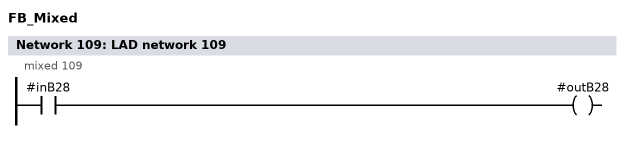
   RUNG wire#powerrail
      Contact( #inB28 )
      Coil( #outB28 )
   END_RUNG
   // the same network as SCL:
   #outB28 := #inB28;
END_REGION

REGION Network 110 (FBD): FBD network 110
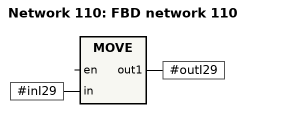
   #outI29 := #inI29;
END_REGION

REGION Network 111 (SCL): SCL network 111
   #tI10 := #inI30 + #cI20;
           IF #inB30 THEN
               #outR10 := #inR10 * 2.0;
           END_IF;
END_REGION

REGION Network 112: LAD network 112
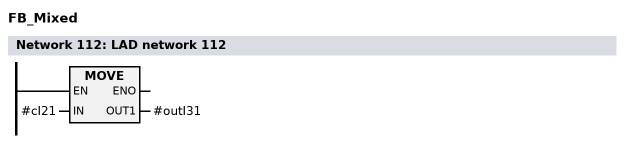
   RUNG wire#powerrail
      Move(in := #cI21, out1 => #outI31)
   END_RUNG
   // the same network as SCL:
   #outI31 := #cI21;
END_REGION

REGION Network 113 (FBD): FBD network 113
   // mixed 113
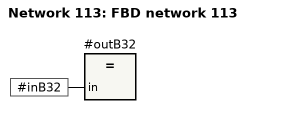
   #outB32 := #inB32;
END_REGION

REGION Network 114 (SCL): SCL network 114
   #tI13 := #inI33 + #cI23;
           IF #inB33 THEN
               #outR13 := #inR13 * 2.0;
           END_IF;
END_REGION

REGION Network 115: LAD network 115
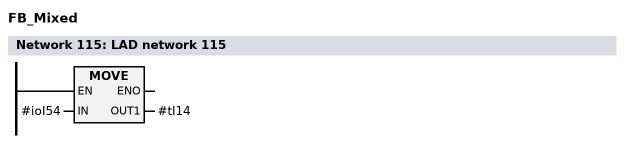
   RUNG wire#powerrail
      Move(in := #ioI54, out1 => #tI14)
   END_RUNG
   // the same network as SCL:
   #tI14 := #ioI54;
END_REGION

REGION Network 116 (FBD): FBD network 116
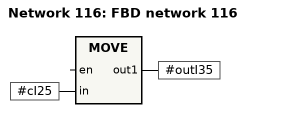
   #outI35 := #cI25;
END_REGION

REGION Network 117 (SCL): SCL network 117
   // mixed 117
   #tI16 := #inI36 + #cI26;
           IF #inB36 THEN
               #outR16 := #inR16 * 2.0;
           END_IF;
END_REGION

REGION Network 118: LAD network 118
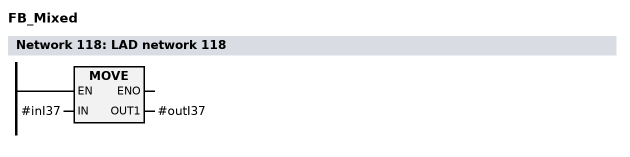
   RUNG wire#powerrail
      Move(in := #inI37, out1 => #outI37)
   END_RUNG
   // the same network as SCL:
   #outI37 := #inI37;
END_REGION

REGION Network 119 (FBD): FBD network 119
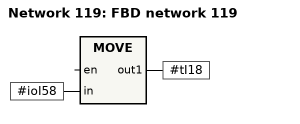
   #tI18 := #ioI58;
END_REGION

REGION Network 120 (SCL): SCL network 120
   #tI19 := #inI39 + #cI29;
           IF #inB39 THEN
               #outR19 := #inR19 * 2.0;
           END_IF;
END_REGION
END_FUNCTION_BLOCK

FUNCTION_BLOCK "FB_BigLad"   // FB14, LAD
{ S7_Optimized_Access := 'TRUE' }
VERSION : 0.1
   VAR_INPUT
      inB0 : Bool;   // input bit 0
      inB1 : Bool;
      inB2 : Bool;
      inB3 : Bool;
      inB4 : Bool;
      inB5 : Bool;
      inB6 : Bool;
      inB7 : Bool;
      inB8 : Bool;
      inB9 : Bool;
      inB10 : Bool;   // input bit 10
      inB11 : Bool;
      inB12 : Bool;
      inB13 : Bool;
      inB14 : Bool;
      inB15 : Bool;
      inB16 : Bool;
      inB17 : Bool;
      inB18 : Bool;
      inB19 : Bool;
      inB20 : Bool;   // input bit 20
      inB21 : Bool;
      inB22 : Bool;
      inB23 : Bool;
      inB24 : Bool;
      inB25 : Bool;
      inB26 : Bool;
      inB27 : Bool;
      inB28 : Bool;
      inB29 : Bool;
      inB30 : Bool;   // input bit 30
      inB31 : Bool;
      inB32 : Bool;
      inB33 : Bool;
      inB34 : Bool;
      inB35 : Bool;
      inB36 : Bool;
      inB37 : Bool;
      inB38 : Bool;
      inB39 : Bool;
      inI0 : Int;
      inI1 : Int;
      inI2 : Int;
      inI3 : Int;
      inI4 : Int;
      inI5 : Int;
      inI6 : Int;
      inI7 : Int;
      inI8 : Int;
      inI9 : Int;
      inI10 : Int;
      inI11 : Int;
      inI12 : Int;
      inI13 : Int;
      inI14 : Int;
      inI15 : Int;
      inI16 : Int;
      inI17 : Int;
      inI18 : Int;
      inI19 : Int;
      inI20 : Int;
      inI21 : Int;
      inI22 : Int;
      inI23 : Int;
      inI24 : Int;
      inI25 : Int;
      inI26 : Int;
      inI27 : Int;
      inI28 : Int;
      inI29 : Int;
      inI30 : Int;
      inI31 : Int;
      inI32 : Int;
      inI33 : Int;
      inI34 : Int;
      inI35 : Int;
      inI36 : Int;
      inI37 : Int;
      inI38 : Int;
      inI39 : Int;
      inR0 : Real;
      inR1 : Real;
      inR2 : Real;
      inR3 : Real;
      inR4 : Real;
      inR5 : Real;
      inR6 : Real;
      inR7 : Real;
      inR8 : Real;
      inR9 : Real;
      inR10 : Real;
      inR11 : Real;
      inR12 : Real;
      inR13 : Real;
      inR14 : Real;
      inR15 : Real;
      inR16 : Real;
      inR17 : Real;
      inR18 : Real;
      inR19 : Real;
      inD0 : DInt;
      inD1 : DInt;
      inD2 : DInt;
      inD3 : DInt;
      inD4 : DInt;
      inD5 : DInt;
      inD6 : DInt;
      inD7 : DInt;
      inD8 : DInt;
      inD9 : DInt;
      inD10 : DInt;
      inD11 : DInt;
      inD12 : DInt;
      inD13 : DInt;
      inD14 : DInt;
      inD15 : DInt;
      inD16 : DInt;
      inD17 : DInt;
      inD18 : DInt;
      inD19 : DInt;
      inArr : Array[0..99] of Int;   // input array
      inStr : String[40];
      inSt : Struct
         x : Int;
         y : Real;
         z : Bool;
      END_STRUCT;
   END_VAR
   VAR_OUTPUT
      outB0 : Bool;
      outB1 : Bool;
      outB2 : Bool;
      outB3 : Bool;
      outB4 : Bool;
      outB5 : Bool;
      outB6 : Bool;
      outB7 : Bool;
      outB8 : Bool;
      outB9 : Bool;
      outB10 : Bool;
      outB11 : Bool;
      outB12 : Bool;
      outB13 : Bool;
      outB14 : Bool;
      outB15 : Bool;
      outB16 : Bool;
      outB17 : Bool;
      outB18 : Bool;
      outB19 : Bool;
      outB20 : Bool;
      outB21 : Bool;
      outB22 : Bool;
      outB23 : Bool;
      outB24 : Bool;
      outB25 : Bool;
      outB26 : Bool;
      outB27 : Bool;
      outB28 : Bool;
      outB29 : Bool;
      outB30 : Bool;
      outB31 : Bool;
      outB32 : Bool;
      outB33 : Bool;
      outB34 : Bool;
      outB35 : Bool;
      outB36 : Bool;
      outB37 : Bool;
      outB38 : Bool;
      outB39 : Bool;
      outI0 : Int;   // output int 0
      outI1 : Int;
      outI2 : Int;
      outI3 : Int;
      outI4 : Int;
      outI5 : Int;
      outI6 : Int;
      outI7 : Int;
      outI8 : Int;
      outI9 : Int;
      outI10 : Int;   // output int 10
      outI11 : Int;
      outI12 : Int;
      outI13 : Int;
      outI14 : Int;
      outI15 : Int;
      outI16 : Int;
      outI17 : Int;
      outI18 : Int;
      outI19 : Int;
      outI20 : Int;   // output int 20
      outI21 : Int;
      outI22 : Int;
      outI23 : Int;
      outI24 : Int;
      outI25 : Int;
      outI26 : Int;
      outI27 : Int;
      outI28 : Int;
      outI29 : Int;
      outI30 : Int;   // output int 30
      outI31 : Int;
      outI32 : Int;
      outI33 : Int;
      outI34 : Int;
      outI35 : Int;
      outI36 : Int;
      outI37 : Int;
      outI38 : Int;
      outI39 : Int;
      outR0 : Real;
      outR1 : Real;
      outR2 : Real;
      outR3 : Real;
      outR4 : Real;
      outR5 : Real;
      outR6 : Real;
      outR7 : Real;
      outR8 : Real;
      outR9 : Real;
      outR10 : Real;
      outR11 : Real;
      outR12 : Real;
      outR13 : Real;
      outR14 : Real;
      outR15 : Real;
      outR16 : Real;
      outR17 : Real;
      outR18 : Real;
      outR19 : Real;
      outD0 : DInt;
      outD1 : DInt;
      outD2 : DInt;
      outD3 : DInt;
      outD4 : DInt;
      outD5 : DInt;
      outD6 : DInt;
      outD7 : DInt;
      outD8 : DInt;
      outD9 : DInt;
      outD10 : DInt;
      outD11 : DInt;
      outD12 : DInt;
      outD13 : DInt;
      outD14 : DInt;
      outD15 : DInt;
      outD16 : DInt;
      outD17 : DInt;
      outD18 : DInt;
      outD19 : DInt;
   END_VAR
   VAR_IN_OUT
      ioI0 : Int;
      ioI1 : Int;
      ioI2 : Int;
      ioI3 : Int;
      ioI4 : Int;
      ioI5 : Int;
      ioI6 : Int;
      ioI7 : Int;
      ioI8 : Int;
      ioI9 : Int;
      ioI10 : Int;
      ioI11 : Int;
      ioI12 : Int;
      ioI13 : Int;
      ioI14 : Int;
      ioI15 : Int;
      ioI16 : Int;
      ioI17 : Int;
      ioI18 : Int;
      ioI19 : Int;
      ioI20 : Int;
      ioI21 : Int;
      ioI22 : Int;
      ioI23 : Int;
      ioI24 : Int;
      ioI25 : Int;
      ioI26 : Int;
      ioI27 : Int;
      ioI28 : Int;
      ioI29 : Int;
      ioI30 : Int;
      ioI31 : Int;
      ioI32 : Int;
      ioI33 : Int;
      ioI34 : Int;
      ioI35 : Int;
      ioI36 : Int;
      ioI37 : Int;
      ioI38 : Int;
      ioI39 : Int;
      ioI40 : Int;
      ioI41 : Int;
      ioI42 : Int;
      ioI43 : Int;
      ioI44 : Int;
      ioI45 : Int;
      ioI46 : Int;
      ioI47 : Int;
      ioI48 : Int;
      ioI49 : Int;
      ioI50 : Int;
      ioI51 : Int;
      ioI52 : Int;
      ioI53 : Int;
      ioI54 : Int;
      ioI55 : Int;
      ioI56 : Int;
      ioI57 : Int;
      ioI58 : Int;
      ioI59 : Int;
   END_VAR
   VAR
      stI0 : Int := 0;   // static 0
      stI1 : Int;
      stI2 : Int;
      stI3 : Int;
      stI4 : Int;
      stI5 : Int;
      stI6 : Int;
      stI7 : Int := 7;
      stI8 : Int;
      stI9 : Int;
      stI10 : Int;
      stI11 : Int;
      stI12 : Int;
      stI13 : Int;
      stI14 : Int := 14;
      stI15 : Int;
      stI16 : Int;
      stI17 : Int;
      stI18 : Int;
      stI19 : Int;
      stI20 : Int;
      stI21 : Int := 21;
      stI22 : Int;
      stI23 : Int;
      stI24 : Int;
      stI25 : Int;   // static 25
      stI26 : Int;
      stI27 : Int;
      stI28 : Int := 28;
      stI29 : Int;
      stI30 : Int;
      stI31 : Int;
      stI32 : Int;
      stI33 : Int;
      stI34 : Int;
      stI35 : Int := 35;
      stI36 : Int;
      stI37 : Int;
      stI38 : Int;
      stI39 : Int;
      stI40 : Int;
      stI41 : Int;
      stI42 : Int := 42;
      stI43 : Int;
      stI44 : Int;
      stI45 : Int;
      stI46 : Int;
      stI47 : Int;
      stI48 : Int;
      stI49 : Int := 49;
      stI50 : Int;   // static 50
      stI51 : Int;
      stI52 : Int;
      stI53 : Int;
      stI54 : Int;
      stI55 : Int;
      stI56 : Int := 56;
      stI57 : Int;
      stI58 : Int;
      stI59 : Int;
      stI60 : Int;
      stI61 : Int;
      stI62 : Int;
      stI63 : Int := 63;
      stI64 : Int;
      stI65 : Int;
      stI66 : Int;
      stI67 : Int;
      stI68 : Int;
      stI69 : Int;
      stI70 : Int := 70;
      stI71 : Int;
      stI72 : Int;
      stI73 : Int;
      stI74 : Int;
      stI75 : Int;   // static 75
      stI76 : Int;
      stI77 : Int := 77;
      stI78 : Int;
      stI79 : Int;
      stI80 : Int;
      stI81 : Int;
      stI82 : Int;
      stI83 : Int;
      stI84 : Int := 84;
      stI85 : Int;
      stI86 : Int;
      stI87 : Int;
      stI88 : Int;
      stI89 : Int;
      stI90 : Int;
      stI91 : Int := 91;
      stI92 : Int;
      stI93 : Int;
      stI94 : Int;
      stI95 : Int;
      stI96 : Int;
      stI97 : Int;
      stI98 : Int := 98;
      stI99 : Int;
      stI100 : Int;   // static 100
      stI101 : Int;
      stI102 : Int;
      stI103 : Int;
      stI104 : Int;
      stI105 : Int := 105;
      stI106 : Int;
      stI107 : Int;
      stI108 : Int;
      stI109 : Int;
      stI110 : Int;
      stI111 : Int;
      stI112 : Int := 112;
      stI113 : Int;
      stI114 : Int;
      stI115 : Int;
      stI116 : Int;
      stI117 : Int;
      stI118 : Int;
      stI119 : Int := 119;
      stI120 : Int;
      stI121 : Int;
      stI122 : Int;
      stI123 : Int;
      stI124 : Int;
      stI125 : Int;   // static 125
      stI126 : Int := 126;
      stI127 : Int;
      stI128 : Int;
      stI129 : Int;
      stI130 : Int;
      stI131 : Int;
      stI132 : Int;
      stI133 : Int := 133;
      stI134 : Int;
      stI135 : Int;
      stI136 : Int;
      stI137 : Int;
      stI138 : Int;
      stI139 : Int;
      stI140 : Int := 140;
      stI141 : Int;
      stI142 : Int;
      stI143 : Int;
      stI144 : Int;
      stI145 : Int;
      stI146 : Int;
      stI147 : Int := 147;
      stI148 : Int;
      stI149 : Int;
      stI150 : Int;   // static 150
      stI151 : Int;
      stI152 : Int;
      stI153 : Int;
      stI154 : Int := 154;
      stI155 : Int;
      stI156 : Int;
      stI157 : Int;
      stI158 : Int;
      stI159 : Int;
      stI160 : Int;
      stI161 : Int := 161;
      stI162 : Int;
      stI163 : Int;
      stI164 : Int;
      stI165 : Int;
      stI166 : Int;
      stI167 : Int;
      stI168 : Int := 168;
      stI169 : Int;
      stI170 : Int;
      stI171 : Int;
      stI172 : Int;
      stI173 : Int;
      stI174 : Int;
      stI175 : Int := 175;   // static 175
      stI176 : Int;
      stI177 : Int;
      stI178 : Int;
      stI179 : Int;
      stI180 : Int;
      stI181 : Int;
      stI182 : Int := 182;
      stI183 : Int;
      stI184 : Int;
      stI185 : Int;
      stI186 : Int;
      stI187 : Int;
      stI188 : Int;
      stI189 : Int := 189;
      stI190 : Int;
      stI191 : Int;
      stI192 : Int;
      stI193 : Int;
      stI194 : Int;
      stI195 : Int;
      stI196 : Int := 196;
      stI197 : Int;
      stI198 : Int;
      stI199 : Int;
      stB0 : Bool := TRUE;
      stB1 : Bool;
      stB2 : Bool;
      stB3 : Bool := TRUE;
      stB4 : Bool;
      stB5 : Bool;
      stB6 : Bool := TRUE;
      stB7 : Bool;
      stB8 : Bool;
      stB9 : Bool := TRUE;
      stB10 : Bool;
      stB11 : Bool;
      stB12 : Bool := TRUE;
      stB13 : Bool;
      stB14 : Bool;
      stB15 : Bool := TRUE;
      stB16 : Bool;
      stB17 : Bool;
      stB18 : Bool := TRUE;
      stB19 : Bool;
      stB20 : Bool;
      stB21 : Bool := TRUE;
      stB22 : Bool;
      stB23 : Bool;
      stB24 : Bool := TRUE;
      stB25 : Bool;
      stB26 : Bool;
      stB27 : Bool := TRUE;
      stB28 : Bool;
      stB29 : Bool;
      stB30 : Bool := TRUE;
      stB31 : Bool;
      stB32 : Bool;
      stB33 : Bool := TRUE;
      stB34 : Bool;
      stB35 : Bool;
      stB36 : Bool := TRUE;
      stB37 : Bool;
      stB38 : Bool;
      stB39 : Bool := TRUE;
      stB40 : Bool;
      stB41 : Bool;
      stB42 : Bool := TRUE;
      stB43 : Bool;
      stB44 : Bool;
      stB45 : Bool := TRUE;
      stB46 : Bool;
      stB47 : Bool;
      stB48 : Bool := TRUE;
      stB49 : Bool;
      stB50 : Bool;
      stB51 : Bool := TRUE;
      stB52 : Bool;
      stB53 : Bool;
      stB54 : Bool := TRUE;
      stB55 : Bool;
      stB56 : Bool;
      stB57 : Bool := TRUE;
      stB58 : Bool;
      stB59 : Bool;
      stB60 : Bool := TRUE;
      stB61 : Bool;
      stB62 : Bool;
      stB63 : Bool := TRUE;
      stB64 : Bool;
      stB65 : Bool;
      stB66 : Bool := TRUE;
      stB67 : Bool;
      stB68 : Bool;
      stB69 : Bool := TRUE;
      stB70 : Bool;
      stB71 : Bool;
      stB72 : Bool := TRUE;
      stB73 : Bool;
      stB74 : Bool;
      stB75 : Bool := TRUE;
      stB76 : Bool;
      stB77 : Bool;
      stB78 : Bool := TRUE;
      stB79 : Bool;
      stB80 : Bool;
      stB81 : Bool := TRUE;
      stB82 : Bool;
      stB83 : Bool;
      stB84 : Bool := TRUE;
      stB85 : Bool;
      stB86 : Bool;
      stB87 : Bool := TRUE;
      stB88 : Bool;
      stB89 : Bool;
      stB90 : Bool := TRUE;
      stB91 : Bool;
      stB92 : Bool;
      stB93 : Bool := TRUE;
      stB94 : Bool;
      stB95 : Bool;
      stB96 : Bool := TRUE;
      stB97 : Bool;
      stB98 : Bool;
      stB99 : Bool := TRUE;
      stArr : Array[1..10, 0..4] of Real;
      stSt : Struct
         "a" : Int;
         "b" : Array[0..3] of Bool;
         c : Time;
      END_STRUCT;
   END_VAR
   VAR_TEMP
      tI0 : Int;
      tI1 : Int;
      tI2 : Int;
      tI3 : Int;
      tI4 : Int;
      tI5 : Int;
      tI6 : Int;
      tI7 : Int;
      tI8 : Int;
      tI9 : Int;
      tI10 : Int;
      tI11 : Int;
      tI12 : Int;
      tI13 : Int;
      tI14 : Int;
      tI15 : Int;
      tI16 : Int;
      tI17 : Int;
      tI18 : Int;
      tI19 : Int;
      tI20 : Int;
      tI21 : Int;
      tI22 : Int;
      tI23 : Int;
      tI24 : Int;
      tI25 : Int;
      tI26 : Int;
      tI27 : Int;
      tI28 : Int;
      tI29 : Int;
      tI30 : Int;
      tI31 : Int;
      tI32 : Int;
      tI33 : Int;
      tI34 : Int;
      tI35 : Int;
      tI36 : Int;
      tI37 : Int;
      tI38 : Int;
      tI39 : Int;
      tI40 : Int;
      tI41 : Int;
      tI42 : Int;
      tI43 : Int;
      tI44 : Int;
      tI45 : Int;
      tI46 : Int;
      tI47 : Int;
      tI48 : Int;
      tI49 : Int;
      tI50 : Int;
      tI51 : Int;
      tI52 : Int;
      tI53 : Int;
      tI54 : Int;
      tI55 : Int;
      tI56 : Int;
      tI57 : Int;
      tI58 : Int;
      tI59 : Int;
      tI60 : Int;
      tI61 : Int;
      tI62 : Int;
      tI63 : Int;
      tI64 : Int;
      tI65 : Int;
      tI66 : Int;
      tI67 : Int;
      tI68 : Int;
      tI69 : Int;
      tI70 : Int;
      tI71 : Int;
      tI72 : Int;
      tI73 : Int;
      tI74 : Int;
      tI75 : Int;
      tI76 : Int;
      tI77 : Int;
      tI78 : Int;
      tI79 : Int;
      tI80 : Int;
      tI81 : Int;
      tI82 : Int;
      tI83 : Int;
      tI84 : Int;
      tI85 : Int;
      tI86 : Int;
      tI87 : Int;
      tI88 : Int;
      tI89 : Int;
      tI90 : Int;
      tI91 : Int;
      tI92 : Int;
      tI93 : Int;
      tI94 : Int;
      tI95 : Int;
      tI96 : Int;
      tI97 : Int;
      tI98 : Int;
      tI99 : Int;
      tR0 : Real;
      tR1 : Real;
      tR2 : Real;
      tR3 : Real;
      tR4 : Real;
      tR5 : Real;
      tR6 : Real;
      tR7 : Real;
      tR8 : Real;
      tR9 : Real;
      tR10 : Real;
      tR11 : Real;
      tR12 : Real;
      tR13 : Real;
      tR14 : Real;
      tR15 : Real;
      tR16 : Real;
      tR17 : Real;
      tR18 : Real;
      tR19 : Real;
      tR20 : Real;
      tR21 : Real;
      tR22 : Real;
      tR23 : Real;
      tR24 : Real;
      tR25 : Real;
      tR26 : Real;
      tR27 : Real;
      tR28 : Real;
      tR29 : Real;
      tR30 : Real;
      tR31 : Real;
      tR32 : Real;
      tR33 : Real;
      tR34 : Real;
      tR35 : Real;
      tR36 : Real;
      tR37 : Real;
      tR38 : Real;
      tR39 : Real;
      tR40 : Real;
      tR41 : Real;
      tR42 : Real;
      tR43 : Real;
      tR44 : Real;
      tR45 : Real;
      tR46 : Real;
      tR47 : Real;
      tR48 : Real;
      tR49 : Real;
   END_VAR
   VAR CONSTANT
      cI0 : Int := 0;
      cI1 : Int := 3;
      cI2 : Int := 6;
      cI3 : Int := 9;
      cI4 : Int := 12;
      cI5 : Int := 15;
      cI6 : Int := 18;
      cI7 : Int := 21;
      cI8 : Int := 24;
      cI9 : Int := 27;
      cI10 : Int := 30;
      cI11 : Int := 33;
      cI12 : Int := 36;
      cI13 : Int := 39;
      cI14 : Int := 42;
      cI15 : Int := 45;
      cI16 : Int := 48;
      cI17 : Int := 51;
      cI18 : Int := 54;
      cI19 : Int := 57;
      cI20 : Int := 60;
      cI21 : Int := 63;
      cI22 : Int := 66;
      cI23 : Int := 69;
      cI24 : Int := 72;
      cI25 : Int := 75;
      cI26 : Int := 78;
      cI27 : Int := 81;
      cI28 : Int := 84;
      cI29 : Int := 87;
   END_VAR
BEGIN

REGION Network 1: LAD network 1
   // comment of network 1
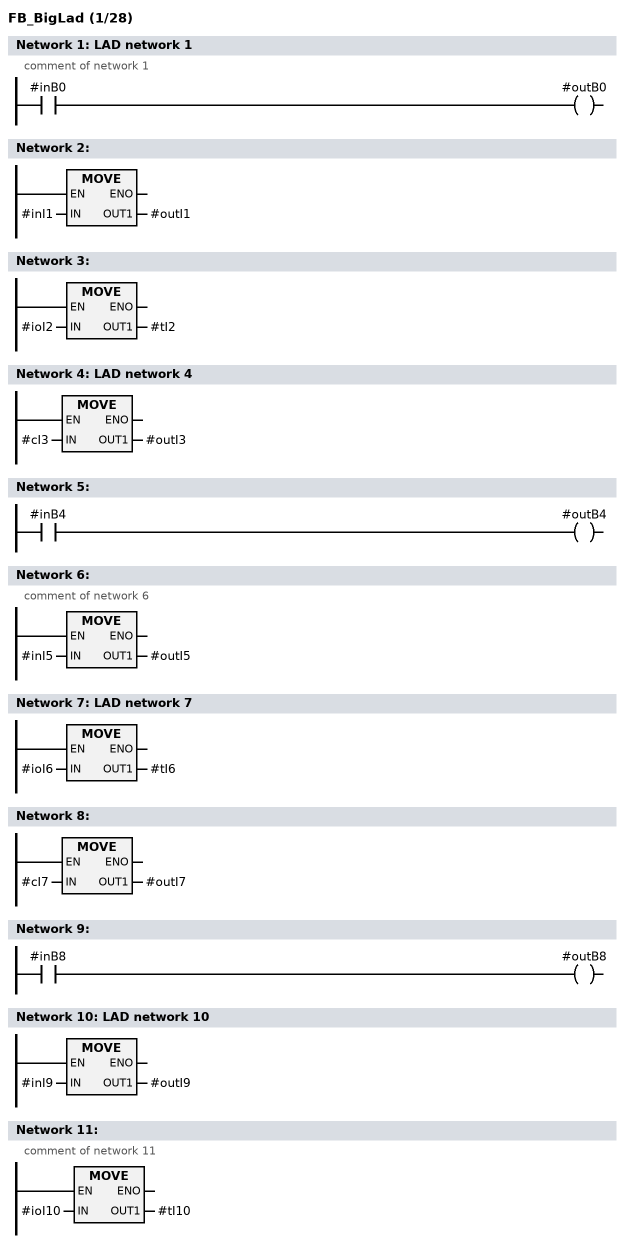
   RUNG wire#powerrail
      Contact( #inB0 )
      Coil( #outB0 )
   END_RUNG
   // the same network as SCL:
   #outB0 := #inB0;
END_REGION

REGION Network 2
   RUNG wire#powerrail
      Move(in := #inI1, out1 => #outI1)
   END_RUNG
   // the same network as SCL:
   #outI1 := #inI1;
END_REGION

REGION Network 3
   RUNG wire#powerrail
      Move(in := #ioI2, out1 => #tI2)
   END_RUNG
   // the same network as SCL:
   #tI2 := #ioI2;
END_REGION

REGION Network 4: LAD network 4
   RUNG wire#powerrail
      Move(in := #cI3, out1 => #outI3)
   END_RUNG
   // the same network as SCL:
   #outI3 := #cI3;
END_REGION

REGION Network 5
   RUNG wire#powerrail
      Contact( #inB4 )
      Coil( #outB4 )
   END_RUNG
   // the same network as SCL:
   #outB4 := #inB4;
END_REGION

REGION Network 6
   // comment of network 6
   RUNG wire#powerrail
      Move(in := #inI5, out1 => #outI5)
   END_RUNG
   // the same network as SCL:
   #outI5 := #inI5;
END_REGION

REGION Network 7: LAD network 7
   RUNG wire#powerrail
      Move(in := #ioI6, out1 => #tI6)
   END_RUNG
   // the same network as SCL:
   #tI6 := #ioI6;
END_REGION

REGION Network 8
   RUNG wire#powerrail
      Move(in := #cI7, out1 => #outI7)
   END_RUNG
   // the same network as SCL:
   #outI7 := #cI7;
END_REGION

REGION Network 9
   RUNG wire#powerrail
      Contact( #inB8 )
      Coil( #outB8 )
   END_RUNG
   // the same network as SCL:
   #outB8 := #inB8;
END_REGION

REGION Network 10: LAD network 10
   RUNG wire#powerrail
      Move(in := #inI9, out1 => #outI9)
   END_RUNG
   // the same network as SCL:
   #outI9 := #inI9;
END_REGION

REGION Network 11
   // comment of network 11
   RUNG wire#powerrail
      Move(in := #ioI10, out1 => #tI10)
   END_RUNG
   // the same network as SCL:
   #tI10 := #ioI10;
END_REGION

REGION Network 12
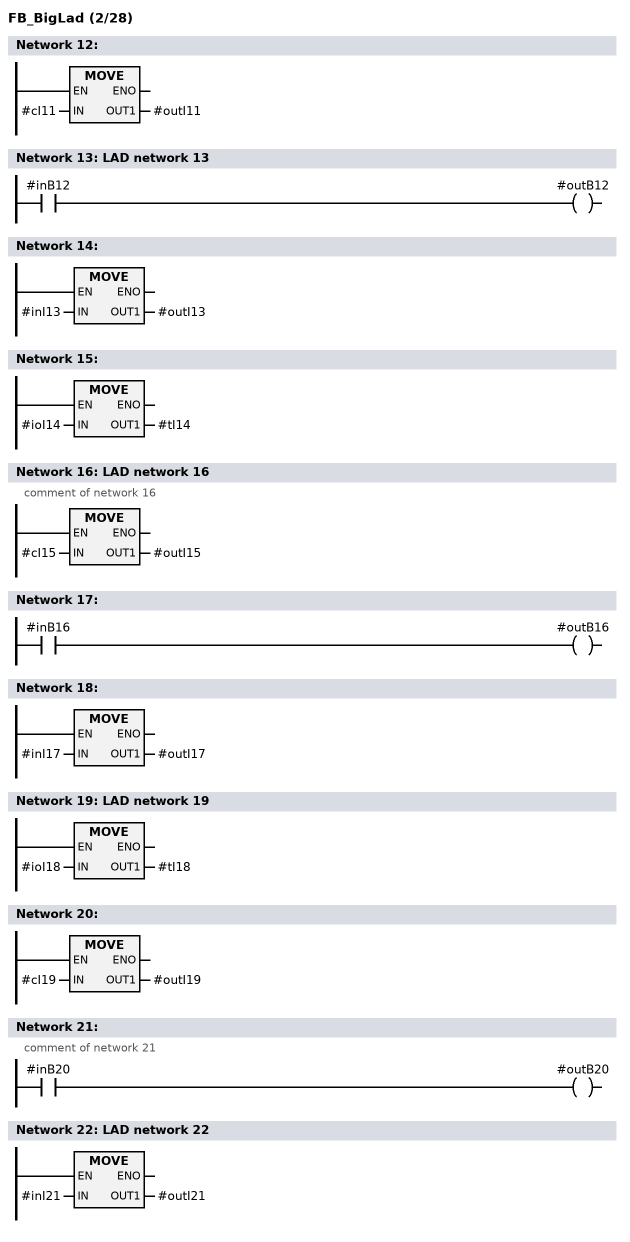
   RUNG wire#powerrail
      Move(in := #cI11, out1 => #outI11)
   END_RUNG
   // the same network as SCL:
   #outI11 := #cI11;
END_REGION

REGION Network 13: LAD network 13
   RUNG wire#powerrail
      Contact( #inB12 )
      Coil( #outB12 )
   END_RUNG
   // the same network as SCL:
   #outB12 := #inB12;
END_REGION

REGION Network 14
   RUNG wire#powerrail
      Move(in := #inI13, out1 => #outI13)
   END_RUNG
   // the same network as SCL:
   #outI13 := #inI13;
END_REGION

REGION Network 15
   RUNG wire#powerrail
      Move(in := #ioI14, out1 => #tI14)
   END_RUNG
   // the same network as SCL:
   #tI14 := #ioI14;
END_REGION

REGION Network 16: LAD network 16
   // comment of network 16
   RUNG wire#powerrail
      Move(in := #cI15, out1 => #outI15)
   END_RUNG
   // the same network as SCL:
   #outI15 := #cI15;
END_REGION

REGION Network 17
   RUNG wire#powerrail
      Contact( #inB16 )
      Coil( #outB16 )
   END_RUNG
   // the same network as SCL:
   #outB16 := #inB16;
END_REGION

REGION Network 18
   RUNG wire#powerrail
      Move(in := #inI17, out1 => #outI17)
   END_RUNG
   // the same network as SCL:
   #outI17 := #inI17;
END_REGION

REGION Network 19: LAD network 19
   RUNG wire#powerrail
      Move(in := #ioI18, out1 => #tI18)
   END_RUNG
   // the same network as SCL:
   #tI18 := #ioI18;
END_REGION

REGION Network 20
   RUNG wire#powerrail
      Move(in := #cI19, out1 => #outI19)
   END_RUNG
   // the same network as SCL:
   #outI19 := #cI19;
END_REGION

REGION Network 21
   // comment of network 21
   RUNG wire#powerrail
      Contact( #inB20 )
      Coil( #outB20 )
   END_RUNG
   // the same network as SCL:
   #outB20 := #inB20;
END_REGION

REGION Network 22: LAD network 22
   RUNG wire#powerrail
      Move(in := #inI21, out1 => #outI21)
   END_RUNG
   // the same network as SCL:
   #outI21 := #inI21;
END_REGION

REGION Network 23
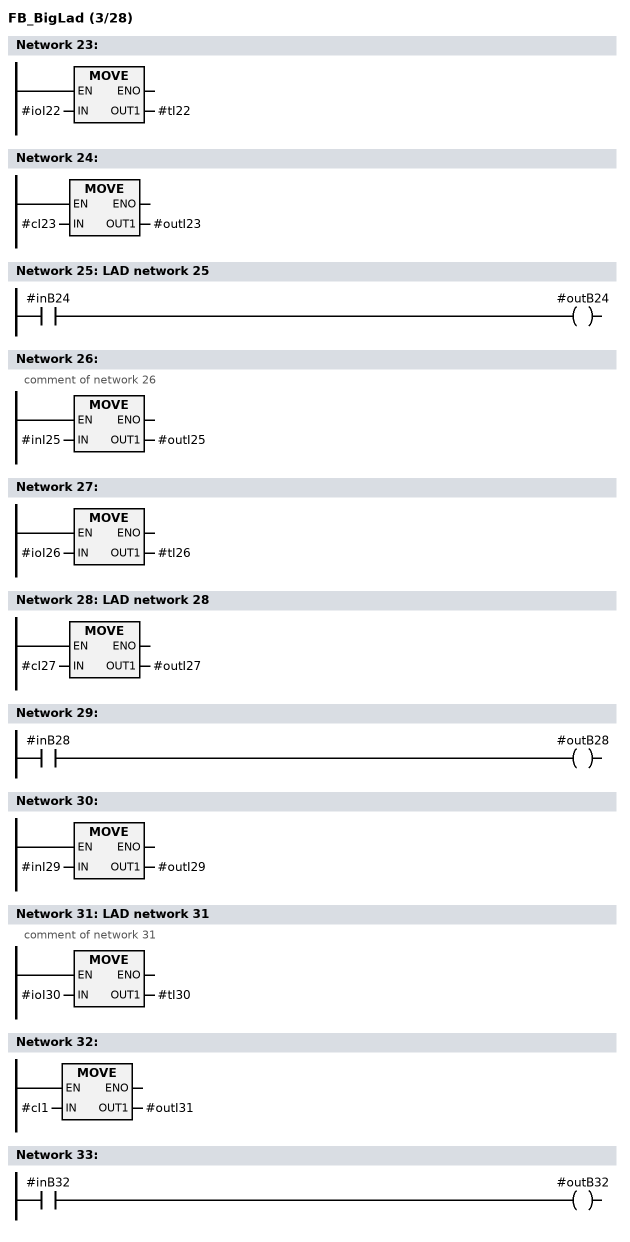
   RUNG wire#powerrail
      Move(in := #ioI22, out1 => #tI22)
   END_RUNG
   // the same network as SCL:
   #tI22 := #ioI22;
END_REGION

REGION Network 24
   RUNG wire#powerrail
      Move(in := #cI23, out1 => #outI23)
   END_RUNG
   // the same network as SCL:
   #outI23 := #cI23;
END_REGION

REGION Network 25: LAD network 25
   RUNG wire#powerrail
      Contact( #inB24 )
      Coil( #outB24 )
   END_RUNG
   // the same network as SCL:
   #outB24 := #inB24;
END_REGION

REGION Network 26
   // comment of network 26
   RUNG wire#powerrail
      Move(in := #inI25, out1 => #outI25)
   END_RUNG
   // the same network as SCL:
   #outI25 := #inI25;
END_REGION

REGION Network 27
   RUNG wire#powerrail
      Move(in := #ioI26, out1 => #tI26)
   END_RUNG
   // the same network as SCL:
   #tI26 := #ioI26;
END_REGION

REGION Network 28: LAD network 28
   RUNG wire#powerrail
      Move(in := #cI27, out1 => #outI27)
   END_RUNG
   // the same network as SCL:
   #outI27 := #cI27;
END_REGION

REGION Network 29
   RUNG wire#powerrail
      Contact( #inB28 )
      Coil( #outB28 )
   END_RUNG
   // the same network as SCL:
   #outB28 := #inB28;
END_REGION

REGION Network 30
   RUNG wire#powerrail
      Move(in := #inI29, out1 => #outI29)
   END_RUNG
   // the same network as SCL:
   #outI29 := #inI29;
END_REGION

REGION Network 31: LAD network 31
   // comment of network 31
   RUNG wire#powerrail
      Move(in := #ioI30, out1 => #tI30)
   END_RUNG
   // the same network as SCL:
   #tI30 := #ioI30;
END_REGION

REGION Network 32
   RUNG wire#powerrail
      Move(in := #cI1, out1 => #outI31)
   END_RUNG
   // the same network as SCL:
   #outI31 := #cI1;
END_REGION

REGION Network 33
   RUNG wire#powerrail
      Contact( #inB32 )
      Coil( #outB32 )
   END_RUNG
   // the same network as SCL:
   #outB32 := #inB32;
END_REGION

REGION Network 34: LAD network 34
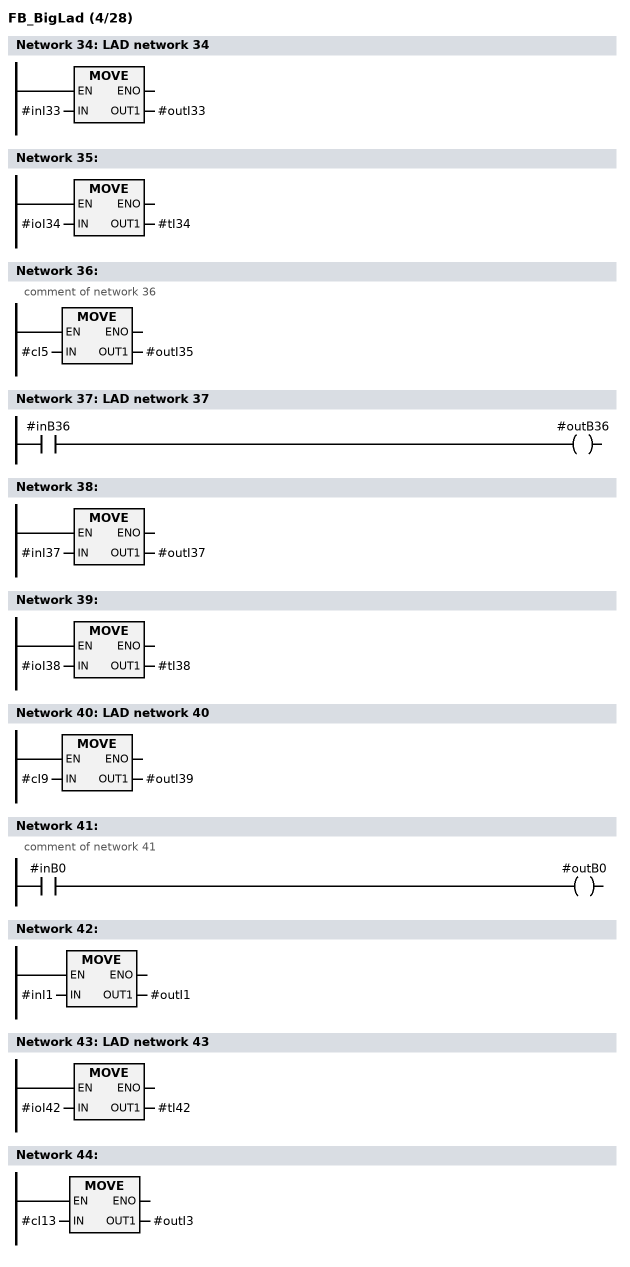
   RUNG wire#powerrail
      Move(in := #inI33, out1 => #outI33)
   END_RUNG
   // the same network as SCL:
   #outI33 := #inI33;
END_REGION

REGION Network 35
   RUNG wire#powerrail
      Move(in := #ioI34, out1 => #tI34)
   END_RUNG
   // the same network as SCL:
   #tI34 := #ioI34;
END_REGION

REGION Network 36
   // comment of network 36
   RUNG wire#powerrail
      Move(in := #cI5, out1 => #outI35)
   END_RUNG
   // the same network as SCL:
   #outI35 := #cI5;
END_REGION

REGION Network 37: LAD network 37
   RUNG wire#powerrail
      Contact( #inB36 )
      Coil( #outB36 )
   END_RUNG
   // the same network as SCL:
   #outB36 := #inB36;
END_REGION

REGION Network 38
   RUNG wire#powerrail
      Move(in := #inI37, out1 => #outI37)
   END_RUNG
   // the same network as SCL:
   #outI37 := #inI37;
END_REGION

REGION Network 39
   RUNG wire#powerrail
      Move(in := #ioI38, out1 => #tI38)
   END_RUNG
   // the same network as SCL:
   #tI38 := #ioI38;
END_REGION

REGION Network 40: LAD network 40
   RUNG wire#powerrail
      Move(in := #cI9, out1 => #outI39)
   END_RUNG
   // the same network as SCL:
   #outI39 := #cI9;
END_REGION

REGION Network 41
   // comment of network 41
   RUNG wire#powerrail
      Contact( #inB0 )
      Coil( #outB0 )
   END_RUNG
   // the same network as SCL:
   #outB0 := #inB0;
END_REGION

REGION Network 42
   RUNG wire#powerrail
      Move(in := #inI1, out1 => #outI1)
   END_RUNG
   // the same network as SCL:
   #outI1 := #inI1;
END_REGION

REGION Network 43: LAD network 43
   RUNG wire#powerrail
      Move(in := #ioI42, out1 => #tI42)
   END_RUNG
   // the same network as SCL:
   #tI42 := #ioI42;
END_REGION

REGION Network 44
   RUNG wire#powerrail
      Move(in := #cI13, out1 => #outI3)
   END_RUNG
   // the same network as SCL:
   #outI3 := #cI13;
END_REGION

REGION Network 45
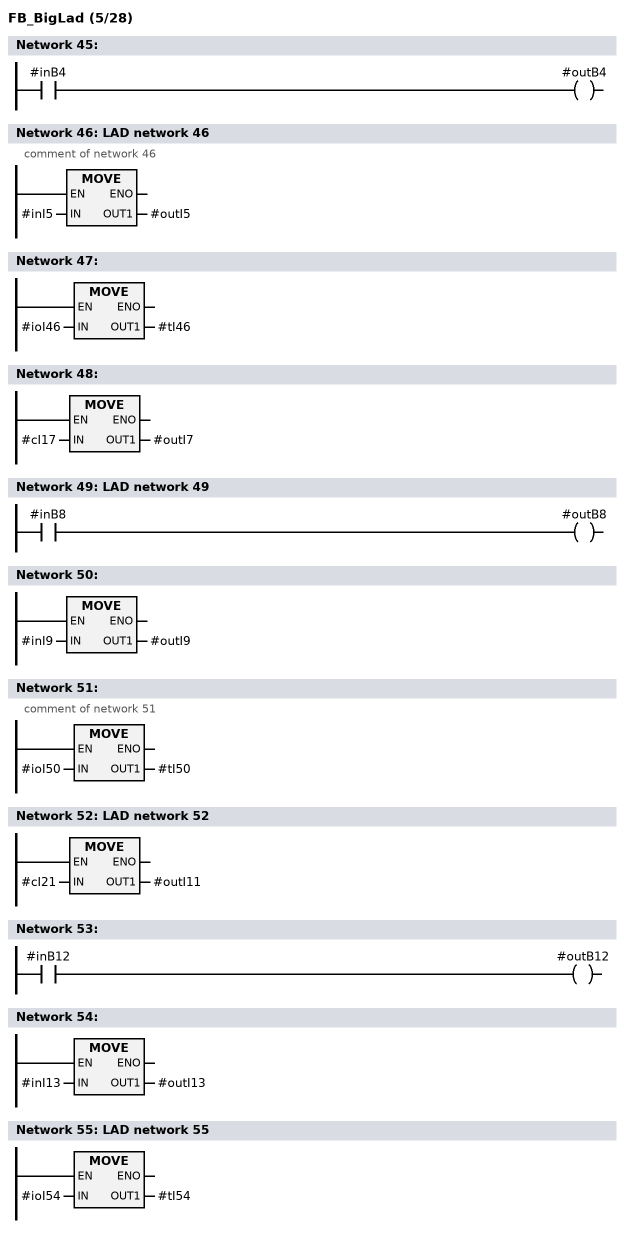
   RUNG wire#powerrail
      Contact( #inB4 )
      Coil( #outB4 )
   END_RUNG
   // the same network as SCL:
   #outB4 := #inB4;
END_REGION

REGION Network 46: LAD network 46
   // comment of network 46
   RUNG wire#powerrail
      Move(in := #inI5, out1 => #outI5)
   END_RUNG
   // the same network as SCL:
   #outI5 := #inI5;
END_REGION

REGION Network 47
   RUNG wire#powerrail
      Move(in := #ioI46, out1 => #tI46)
   END_RUNG
   // the same network as SCL:
   #tI46 := #ioI46;
END_REGION

REGION Network 48
   RUNG wire#powerrail
      Move(in := #cI17, out1 => #outI7)
   END_RUNG
   // the same network as SCL:
   #outI7 := #cI17;
END_REGION

REGION Network 49: LAD network 49
   RUNG wire#powerrail
      Contact( #inB8 )
      Coil( #outB8 )
   END_RUNG
   // the same network as SCL:
   #outB8 := #inB8;
END_REGION

REGION Network 50
   RUNG wire#powerrail
      Move(in := #inI9, out1 => #outI9)
   END_RUNG
   // the same network as SCL:
   #outI9 := #inI9;
END_REGION

REGION Network 51
   // comment of network 51
   RUNG wire#powerrail
      Move(in := #ioI50, out1 => #tI50)
   END_RUNG
   // the same network as SCL:
   #tI50 := #ioI50;
END_REGION

REGION Network 52: LAD network 52
   RUNG wire#powerrail
      Move(in := #cI21, out1 => #outI11)
   END_RUNG
   // the same network as SCL:
   #outI11 := #cI21;
END_REGION

REGION Network 53
   RUNG wire#powerrail
      Contact( #inB12 )
      Coil( #outB12 )
   END_RUNG
   // the same network as SCL:
   #outB12 := #inB12;
END_REGION

REGION Network 54
   RUNG wire#powerrail
      Move(in := #inI13, out1 => #outI13)
   END_RUNG
   // the same network as SCL:
   #outI13 := #inI13;
END_REGION

REGION Network 55: LAD network 55
   RUNG wire#powerrail
      Move(in := #ioI54, out1 => #tI54)
   END_RUNG
   // the same network as SCL:
   #tI54 := #ioI54;
END_REGION

REGION Network 56
   // comment of network 56
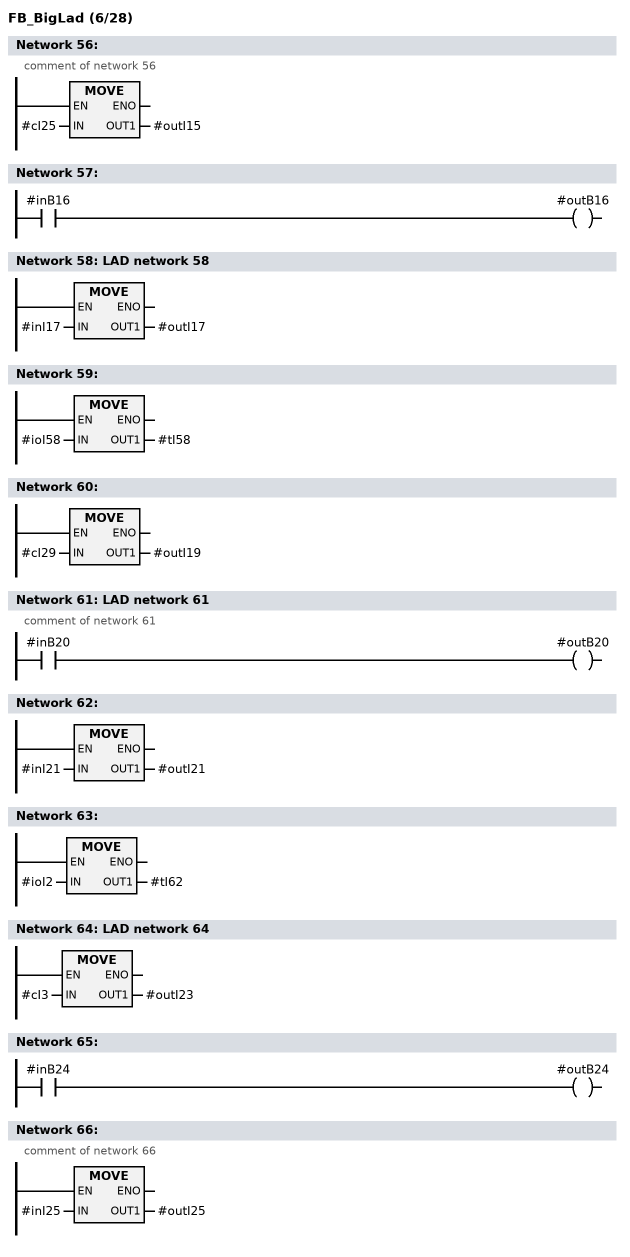
   RUNG wire#powerrail
      Move(in := #cI25, out1 => #outI15)
   END_RUNG
   // the same network as SCL:
   #outI15 := #cI25;
END_REGION

REGION Network 57
   RUNG wire#powerrail
      Contact( #inB16 )
      Coil( #outB16 )
   END_RUNG
   // the same network as SCL:
   #outB16 := #inB16;
END_REGION

REGION Network 58: LAD network 58
   RUNG wire#powerrail
      Move(in := #inI17, out1 => #outI17)
   END_RUNG
   // the same network as SCL:
   #outI17 := #inI17;
END_REGION

REGION Network 59
   RUNG wire#powerrail
      Move(in := #ioI58, out1 => #tI58)
   END_RUNG
   // the same network as SCL:
   #tI58 := #ioI58;
END_REGION

REGION Network 60
   RUNG wire#powerrail
      Move(in := #cI29, out1 => #outI19)
   END_RUNG
   // the same network as SCL:
   #outI19 := #cI29;
END_REGION

REGION Network 61: LAD network 61
   // comment of network 61
   RUNG wire#powerrail
      Contact( #inB20 )
      Coil( #outB20 )
   END_RUNG
   // the same network as SCL:
   #outB20 := #inB20;
END_REGION

REGION Network 62
   RUNG wire#powerrail
      Move(in := #inI21, out1 => #outI21)
   END_RUNG
   // the same network as SCL:
   #outI21 := #inI21;
END_REGION

REGION Network 63
   RUNG wire#powerrail
      Move(in := #ioI2, out1 => #tI62)
   END_RUNG
   // the same network as SCL:
   #tI62 := #ioI2;
END_REGION

REGION Network 64: LAD network 64
   RUNG wire#powerrail
      Move(in := #cI3, out1 => #outI23)
   END_RUNG
   // the same network as SCL:
   #outI23 := #cI3;
END_REGION

REGION Network 65
   RUNG wire#powerrail
      Contact( #inB24 )
      Coil( #outB24 )
   END_RUNG
   // the same network as SCL:
   #outB24 := #inB24;
END_REGION

REGION Network 66
   // comment of network 66
   RUNG wire#powerrail
      Move(in := #inI25, out1 => #outI25)
   END_RUNG
   // the same network as SCL:
   #outI25 := #inI25;
END_REGION

REGION Network 67: LAD network 67
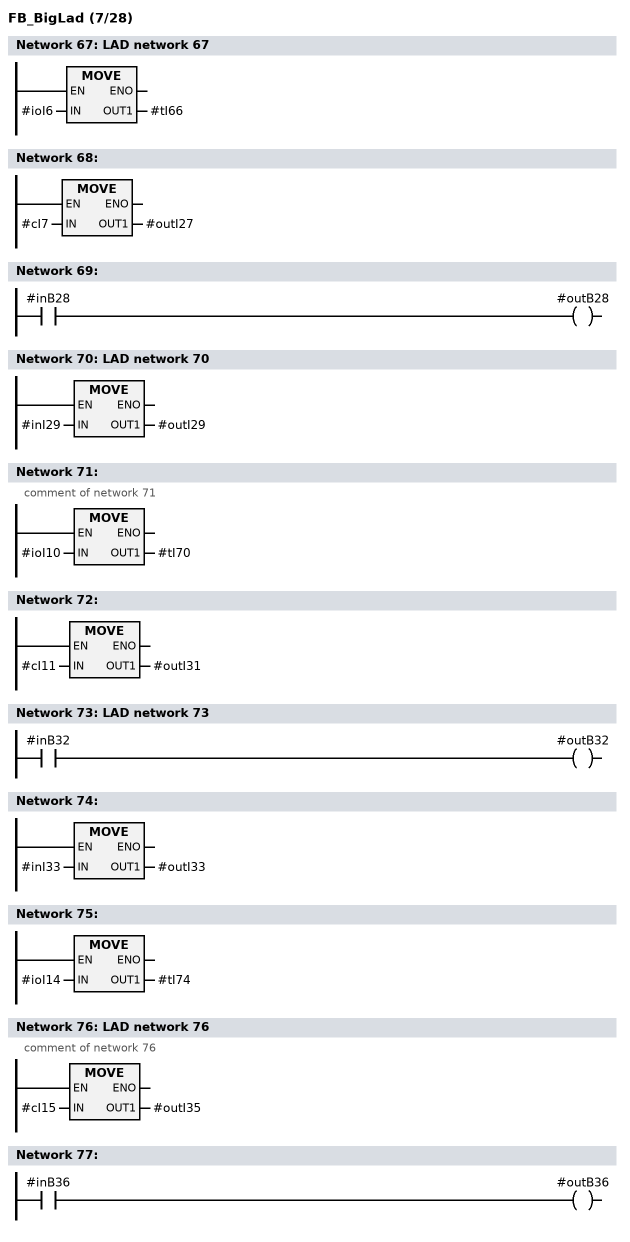
   RUNG wire#powerrail
      Move(in := #ioI6, out1 => #tI66)
   END_RUNG
   // the same network as SCL:
   #tI66 := #ioI6;
END_REGION

REGION Network 68
   RUNG wire#powerrail
      Move(in := #cI7, out1 => #outI27)
   END_RUNG
   // the same network as SCL:
   #outI27 := #cI7;
END_REGION

REGION Network 69
   RUNG wire#powerrail
      Contact( #inB28 )
      Coil( #outB28 )
   END_RUNG
   // the same network as SCL:
   #outB28 := #inB28;
END_REGION

REGION Network 70: LAD network 70
   RUNG wire#powerrail
      Move(in := #inI29, out1 => #outI29)
   END_RUNG
   // the same network as SCL:
   #outI29 := #inI29;
END_REGION

REGION Network 71
   // comment of network 71
   RUNG wire#powerrail
      Move(in := #ioI10, out1 => #tI70)
   END_RUNG
   // the same network as SCL:
   #tI70 := #ioI10;
END_REGION

REGION Network 72
   RUNG wire#powerrail
      Move(in := #cI11, out1 => #outI31)
   END_RUNG
   // the same network as SCL:
   #outI31 := #cI11;
END_REGION

REGION Network 73: LAD network 73
   RUNG wire#powerrail
      Contact( #inB32 )
      Coil( #outB32 )
   END_RUNG
   // the same network as SCL:
   #outB32 := #inB32;
END_REGION

REGION Network 74
   RUNG wire#powerrail
      Move(in := #inI33, out1 => #outI33)
   END_RUNG
   // the same network as SCL:
   #outI33 := #inI33;
END_REGION

REGION Network 75
   RUNG wire#powerrail
      Move(in := #ioI14, out1 => #tI74)
   END_RUNG
   // the same network as SCL:
   #tI74 := #ioI14;
END_REGION

REGION Network 76: LAD network 76
   // comment of network 76
   RUNG wire#powerrail
      Move(in := #cI15, out1 => #outI35)
   END_RUNG
   // the same network as SCL:
   #outI35 := #cI15;
END_REGION

REGION Network 77
   RUNG wire#powerrail
      Contact( #inB36 )
      Coil( #outB36 )
   END_RUNG
   // the same network as SCL:
   #outB36 := #inB36;
END_REGION

REGION Network 78
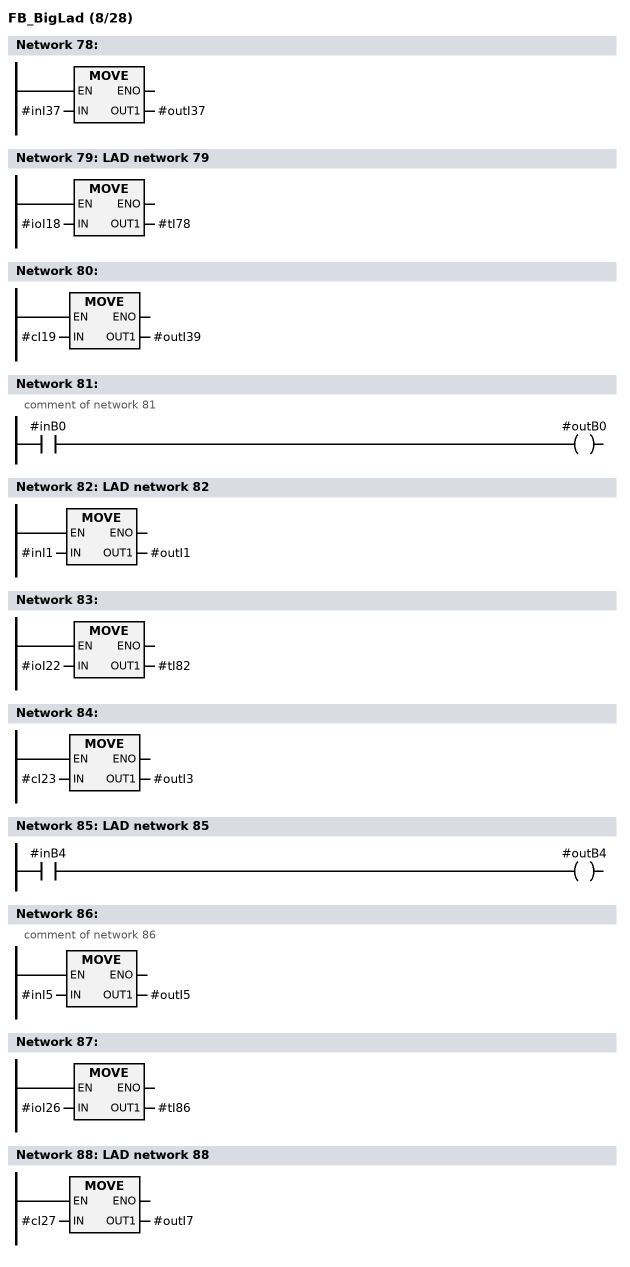
   RUNG wire#powerrail
      Move(in := #inI37, out1 => #outI37)
   END_RUNG
   // the same network as SCL:
   #outI37 := #inI37;
END_REGION

REGION Network 79: LAD network 79
   RUNG wire#powerrail
      Move(in := #ioI18, out1 => #tI78)
   END_RUNG
   // the same network as SCL:
   #tI78 := #ioI18;
END_REGION

REGION Network 80
   RUNG wire#powerrail
      Move(in := #cI19, out1 => #outI39)
   END_RUNG
   // the same network as SCL:
   #outI39 := #cI19;
END_REGION

REGION Network 81
   // comment of network 81
   RUNG wire#powerrail
      Contact( #inB0 )
      Coil( #outB0 )
   END_RUNG
   // the same network as SCL:
   #outB0 := #inB0;
END_REGION

REGION Network 82: LAD network 82
   RUNG wire#powerrail
      Move(in := #inI1, out1 => #outI1)
   END_RUNG
   // the same network as SCL:
   #outI1 := #inI1;
END_REGION

REGION Network 83
   RUNG wire#powerrail
      Move(in := #ioI22, out1 => #tI82)
   END_RUNG
   // the same network as SCL:
   #tI82 := #ioI22;
END_REGION

REGION Network 84
   RUNG wire#powerrail
      Move(in := #cI23, out1 => #outI3)
   END_RUNG
   // the same network as SCL:
   #outI3 := #cI23;
END_REGION

REGION Network 85: LAD network 85
   RUNG wire#powerrail
      Contact( #inB4 )
      Coil( #outB4 )
   END_RUNG
   // the same network as SCL:
   #outB4 := #inB4;
END_REGION

REGION Network 86
   // comment of network 86
   RUNG wire#powerrail
      Move(in := #inI5, out1 => #outI5)
   END_RUNG
   // the same network as SCL:
   #outI5 := #inI5;
END_REGION

REGION Network 87
   RUNG wire#powerrail
      Move(in := #ioI26, out1 => #tI86)
   END_RUNG
   // the same network as SCL:
   #tI86 := #ioI26;
END_REGION

REGION Network 88: LAD network 88
   RUNG wire#powerrail
      Move(in := #cI27, out1 => #outI7)
   END_RUNG
   // the same network as SCL:
   #outI7 := #cI27;
END_REGION

REGION Network 89
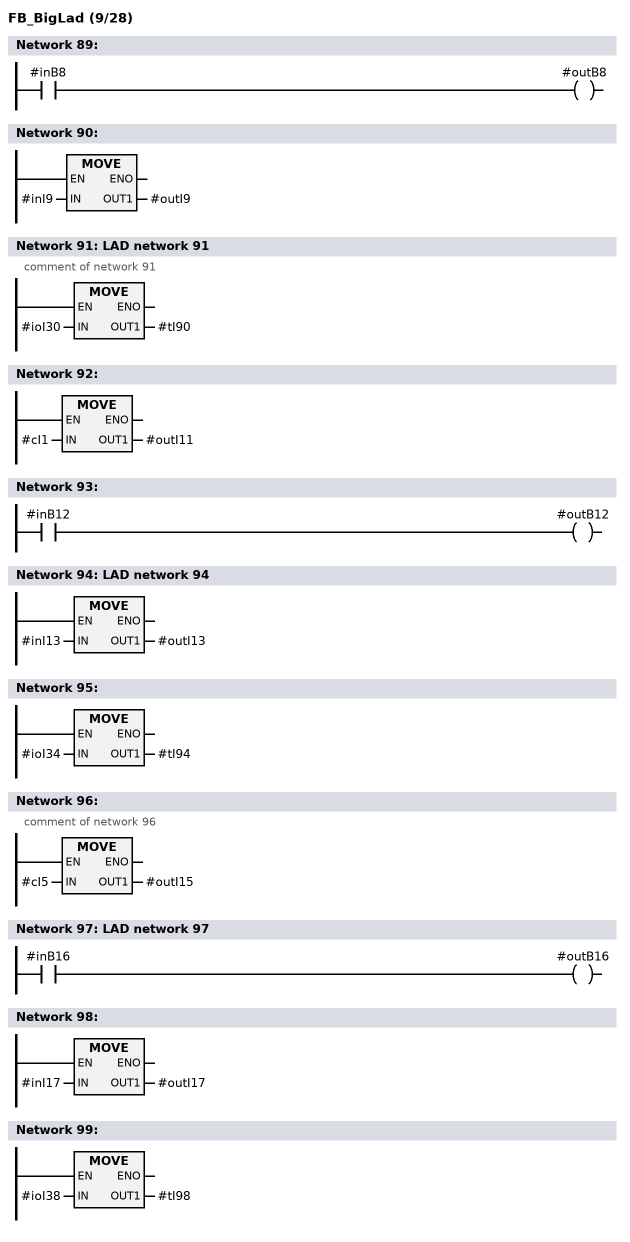
   RUNG wire#powerrail
      Contact( #inB8 )
      Coil( #outB8 )
   END_RUNG
   // the same network as SCL:
   #outB8 := #inB8;
END_REGION

REGION Network 90
   RUNG wire#powerrail
      Move(in := #inI9, out1 => #outI9)
   END_RUNG
   // the same network as SCL:
   #outI9 := #inI9;
END_REGION

REGION Network 91: LAD network 91
   // comment of network 91
   RUNG wire#powerrail
      Move(in := #ioI30, out1 => #tI90)
   END_RUNG
   // the same network as SCL:
   #tI90 := #ioI30;
END_REGION

REGION Network 92
   RUNG wire#powerrail
      Move(in := #cI1, out1 => #outI11)
   END_RUNG
   // the same network as SCL:
   #outI11 := #cI1;
END_REGION

REGION Network 93
   RUNG wire#powerrail
      Contact( #inB12 )
      Coil( #outB12 )
   END_RUNG
   // the same network as SCL:
   #outB12 := #inB12;
END_REGION

REGION Network 94: LAD network 94
   RUNG wire#powerrail
      Move(in := #inI13, out1 => #outI13)
   END_RUNG
   // the same network as SCL:
   #outI13 := #inI13;
END_REGION

REGION Network 95
   RUNG wire#powerrail
      Move(in := #ioI34, out1 => #tI94)
   END_RUNG
   // the same network as SCL:
   #tI94 := #ioI34;
END_REGION

REGION Network 96
   // comment of network 96
   RUNG wire#powerrail
      Move(in := #cI5, out1 => #outI15)
   END_RUNG
   // the same network as SCL:
   #outI15 := #cI5;
END_REGION

REGION Network 97: LAD network 97
   RUNG wire#powerrail
      Contact( #inB16 )
      Coil( #outB16 )
   END_RUNG
   // the same network as SCL:
   #outB16 := #inB16;
END_REGION

REGION Network 98
   RUNG wire#powerrail
      Move(in := #inI17, out1 => #outI17)
   END_RUNG
   // the same network as SCL:
   #outI17 := #inI17;
END_REGION

REGION Network 99
   RUNG wire#powerrail
      Move(in := #ioI38, out1 => #tI98)
   END_RUNG
   // the same network as SCL:
   #tI98 := #ioI38;
END_REGION

REGION Network 100: LAD network 100
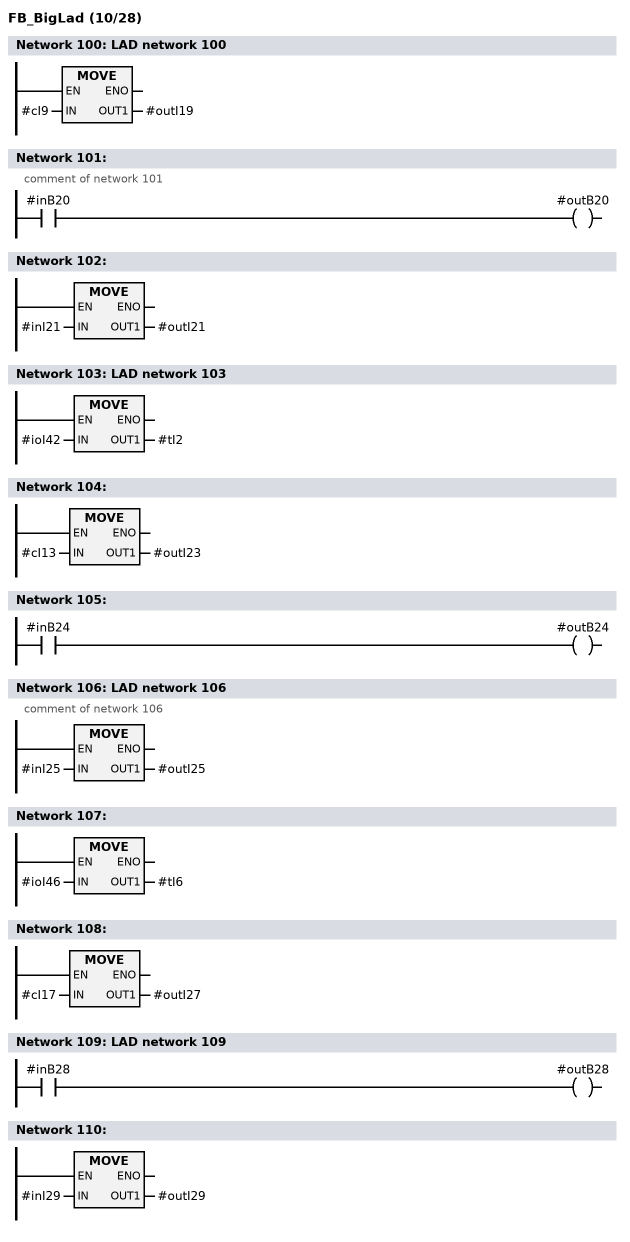
   RUNG wire#powerrail
      Move(in := #cI9, out1 => #outI19)
   END_RUNG
   // the same network as SCL:
   #outI19 := #cI9;
END_REGION

REGION Network 101
   // comment of network 101
   RUNG wire#powerrail
      Contact( #inB20 )
      Coil( #outB20 )
   END_RUNG
   // the same network as SCL:
   #outB20 := #inB20;
END_REGION

REGION Network 102
   RUNG wire#powerrail
      Move(in := #inI21, out1 => #outI21)
   END_RUNG
   // the same network as SCL:
   #outI21 := #inI21;
END_REGION

REGION Network 103: LAD network 103
   RUNG wire#powerrail
      Move(in := #ioI42, out1 => #tI2)
   END_RUNG
   // the same network as SCL:
   #tI2 := #ioI42;
END_REGION

REGION Network 104
   RUNG wire#powerrail
      Move(in := #cI13, out1 => #outI23)
   END_RUNG
   // the same network as SCL:
   #outI23 := #cI13;
END_REGION

REGION Network 105
   RUNG wire#powerrail
      Contact( #inB24 )
      Coil( #outB24 )
   END_RUNG
   // the same network as SCL:
   #outB24 := #inB24;
END_REGION

REGION Network 106: LAD network 106
   // comment of network 106
   RUNG wire#powerrail
      Move(in := #inI25, out1 => #outI25)
   END_RUNG
   // the same network as SCL:
   #outI25 := #inI25;
END_REGION

REGION Network 107
   RUNG wire#powerrail
      Move(in := #ioI46, out1 => #tI6)
   END_RUNG
   // the same network as SCL:
   #tI6 := #ioI46;
END_REGION

REGION Network 108
   RUNG wire#powerrail
      Move(in := #cI17, out1 => #outI27)
   END_RUNG
   // the same network as SCL:
   #outI27 := #cI17;
END_REGION

REGION Network 109: LAD network 109
   RUNG wire#powerrail
      Contact( #inB28 )
      Coil( #outB28 )
   END_RUNG
   // the same network as SCL:
   #outB28 := #inB28;
END_REGION

REGION Network 110
   RUNG wire#powerrail
      Move(in := #inI29, out1 => #outI29)
   END_RUNG
   // the same network as SCL:
   #outI29 := #inI29;
END_REGION

REGION Network 111
   // comment of network 111
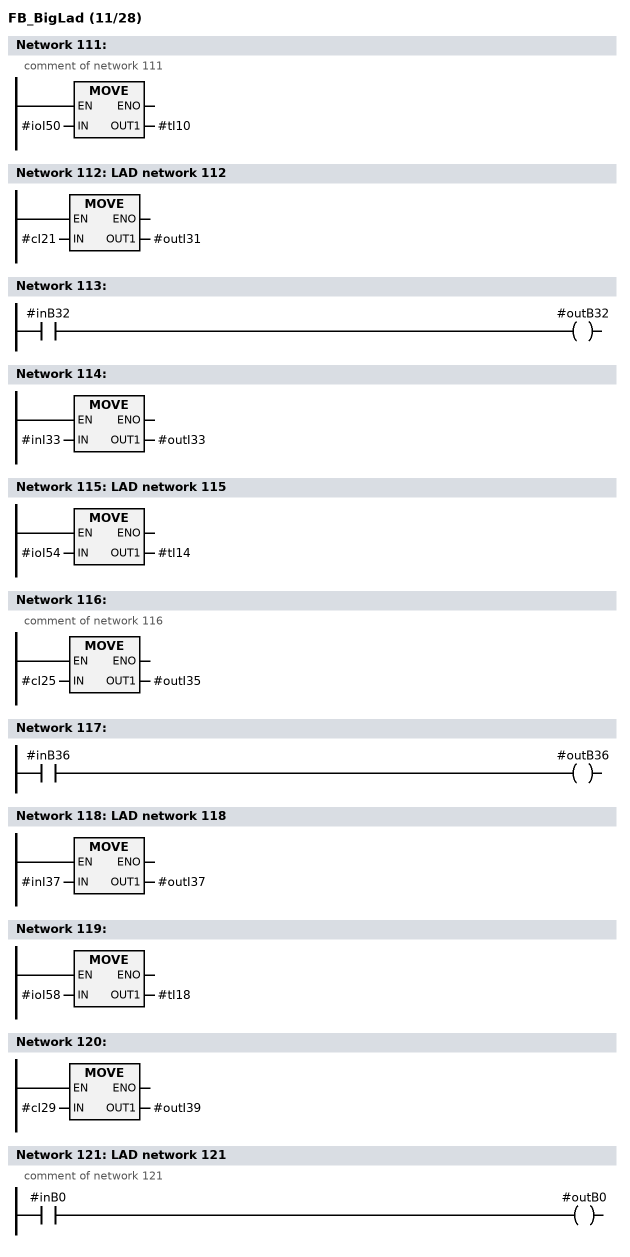
   RUNG wire#powerrail
      Move(in := #ioI50, out1 => #tI10)
   END_RUNG
   // the same network as SCL:
   #tI10 := #ioI50;
END_REGION

REGION Network 112: LAD network 112
   RUNG wire#powerrail
      Move(in := #cI21, out1 => #outI31)
   END_RUNG
   // the same network as SCL:
   #outI31 := #cI21;
END_REGION

REGION Network 113
   RUNG wire#powerrail
      Contact( #inB32 )
      Coil( #outB32 )
   END_RUNG
   // the same network as SCL:
   #outB32 := #inB32;
END_REGION

REGION Network 114
   RUNG wire#powerrail
      Move(in := #inI33, out1 => #outI33)
   END_RUNG
   // the same network as SCL:
   #outI33 := #inI33;
END_REGION

REGION Network 115: LAD network 115
   RUNG wire#powerrail
      Move(in := #ioI54, out1 => #tI14)
   END_RUNG
   // the same network as SCL:
   #tI14 := #ioI54;
END_REGION

REGION Network 116
   // comment of network 116
   RUNG wire#powerrail
      Move(in := #cI25, out1 => #outI35)
   END_RUNG
   // the same network as SCL:
   #outI35 := #cI25;
END_REGION

REGION Network 117
   RUNG wire#powerrail
      Contact( #inB36 )
      Coil( #outB36 )
   END_RUNG
   // the same network as SCL:
   #outB36 := #inB36;
END_REGION

REGION Network 118: LAD network 118
   RUNG wire#powerrail
      Move(in := #inI37, out1 => #outI37)
   END_RUNG
   // the same network as SCL:
   #outI37 := #inI37;
END_REGION

REGION Network 119
   RUNG wire#powerrail
      Move(in := #ioI58, out1 => #tI18)
   END_RUNG
   // the same network as SCL:
   #tI18 := #ioI58;
END_REGION

REGION Network 120
   RUNG wire#powerrail
      Move(in := #cI29, out1 => #outI39)
   END_RUNG
   // the same network as SCL:
   #outI39 := #cI29;
END_REGION

REGION Network 121: LAD network 121
   // comment of network 121
   RUNG wire#powerrail
      Contact( #inB0 )
      Coil( #outB0 )
   END_RUNG
   // the same network as SCL:
   #outB0 := #inB0;
END_REGION

REGION Network 122
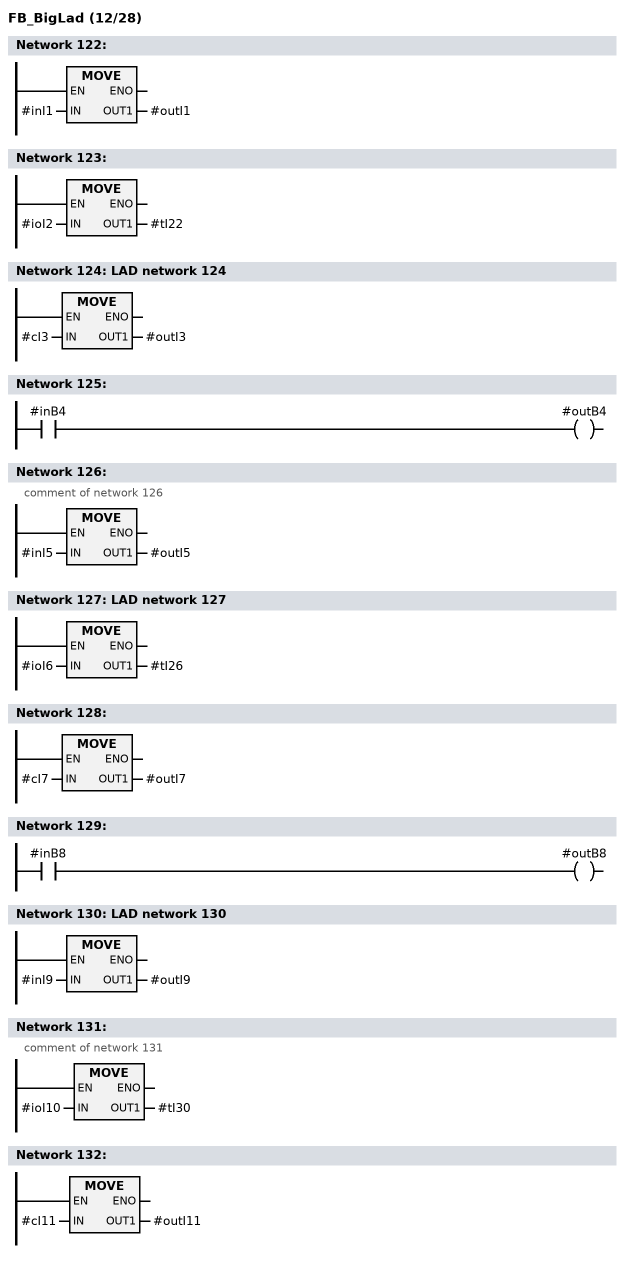
   RUNG wire#powerrail
      Move(in := #inI1, out1 => #outI1)
   END_RUNG
   // the same network as SCL:
   #outI1 := #inI1;
END_REGION

REGION Network 123
   RUNG wire#powerrail
      Move(in := #ioI2, out1 => #tI22)
   END_RUNG
   // the same network as SCL:
   #tI22 := #ioI2;
END_REGION

REGION Network 124: LAD network 124
   RUNG wire#powerrail
      Move(in := #cI3, out1 => #outI3)
   END_RUNG
   // the same network as SCL:
   #outI3 := #cI3;
END_REGION

REGION Network 125
   RUNG wire#powerrail
      Contact( #inB4 )
      Coil( #outB4 )
   END_RUNG
   // the same network as SCL:
   #outB4 := #inB4;
END_REGION

REGION Network 126
   // comment of network 126
   RUNG wire#powerrail
      Move(in := #inI5, out1 => #outI5)
   END_RUNG
   // the same network as SCL:
   #outI5 := #inI5;
END_REGION

REGION Network 127: LAD network 127
   RUNG wire#powerrail
      Move(in := #ioI6, out1 => #tI26)
   END_RUNG
   // the same network as SCL:
   #tI26 := #ioI6;
END_REGION

REGION Network 128
   RUNG wire#powerrail
      Move(in := #cI7, out1 => #outI7)
   END_RUNG
   // the same network as SCL:
   #outI7 := #cI7;
END_REGION

REGION Network 129
   RUNG wire#powerrail
      Contact( #inB8 )
      Coil( #outB8 )
   END_RUNG
   // the same network as SCL:
   #outB8 := #inB8;
END_REGION

REGION Network 130: LAD network 130
   RUNG wire#powerrail
      Move(in := #inI9, out1 => #outI9)
   END_RUNG
   // the same network as SCL:
   #outI9 := #inI9;
END_REGION

REGION Network 131
   // comment of network 131
   RUNG wire#powerrail
      Move(in := #ioI10, out1 => #tI30)
   END_RUNG
   // the same network as SCL:
   #tI30 := #ioI10;
END_REGION

REGION Network 132
   RUNG wire#powerrail
      Move(in := #cI11, out1 => #outI11)
   END_RUNG
   // the same network as SCL:
   #outI11 := #cI11;
END_REGION

REGION Network 133: LAD network 133
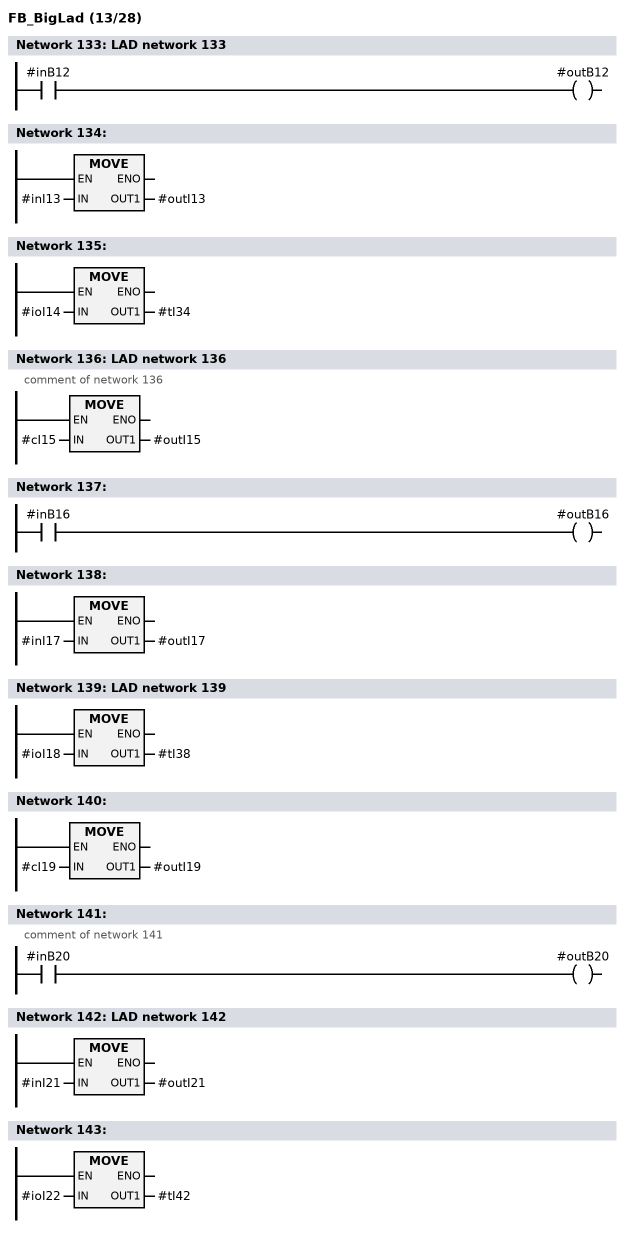
   RUNG wire#powerrail
      Contact( #inB12 )
      Coil( #outB12 )
   END_RUNG
   // the same network as SCL:
   #outB12 := #inB12;
END_REGION

REGION Network 134
   RUNG wire#powerrail
      Move(in := #inI13, out1 => #outI13)
   END_RUNG
   // the same network as SCL:
   #outI13 := #inI13;
END_REGION

REGION Network 135
   RUNG wire#powerrail
      Move(in := #ioI14, out1 => #tI34)
   END_RUNG
   // the same network as SCL:
   #tI34 := #ioI14;
END_REGION

REGION Network 136: LAD network 136
   // comment of network 136
   RUNG wire#powerrail
      Move(in := #cI15, out1 => #outI15)
   END_RUNG
   // the same network as SCL:
   #outI15 := #cI15;
END_REGION

REGION Network 137
   RUNG wire#powerrail
      Contact( #inB16 )
      Coil( #outB16 )
   END_RUNG
   // the same network as SCL:
   #outB16 := #inB16;
END_REGION

REGION Network 138
   RUNG wire#powerrail
      Move(in := #inI17, out1 => #outI17)
   END_RUNG
   // the same network as SCL:
   #outI17 := #inI17;
END_REGION

REGION Network 139: LAD network 139
   RUNG wire#powerrail
      Move(in := #ioI18, out1 => #tI38)
   END_RUNG
   // the same network as SCL:
   #tI38 := #ioI18;
END_REGION

REGION Network 140
   RUNG wire#powerrail
      Move(in := #cI19, out1 => #outI19)
   END_RUNG
   // the same network as SCL:
   #outI19 := #cI19;
END_REGION

REGION Network 141
   // comment of network 141
   RUNG wire#powerrail
      Contact( #inB20 )
      Coil( #outB20 )
   END_RUNG
   // the same network as SCL:
   #outB20 := #inB20;
END_REGION

REGION Network 142: LAD network 142
   RUNG wire#powerrail
      Move(in := #inI21, out1 => #outI21)
   END_RUNG
   // the same network as SCL:
   #outI21 := #inI21;
END_REGION

REGION Network 143
   RUNG wire#powerrail
      Move(in := #ioI22, out1 => #tI42)
   END_RUNG
   // the same network as SCL:
   #tI42 := #ioI22;
END_REGION

REGION Network 144
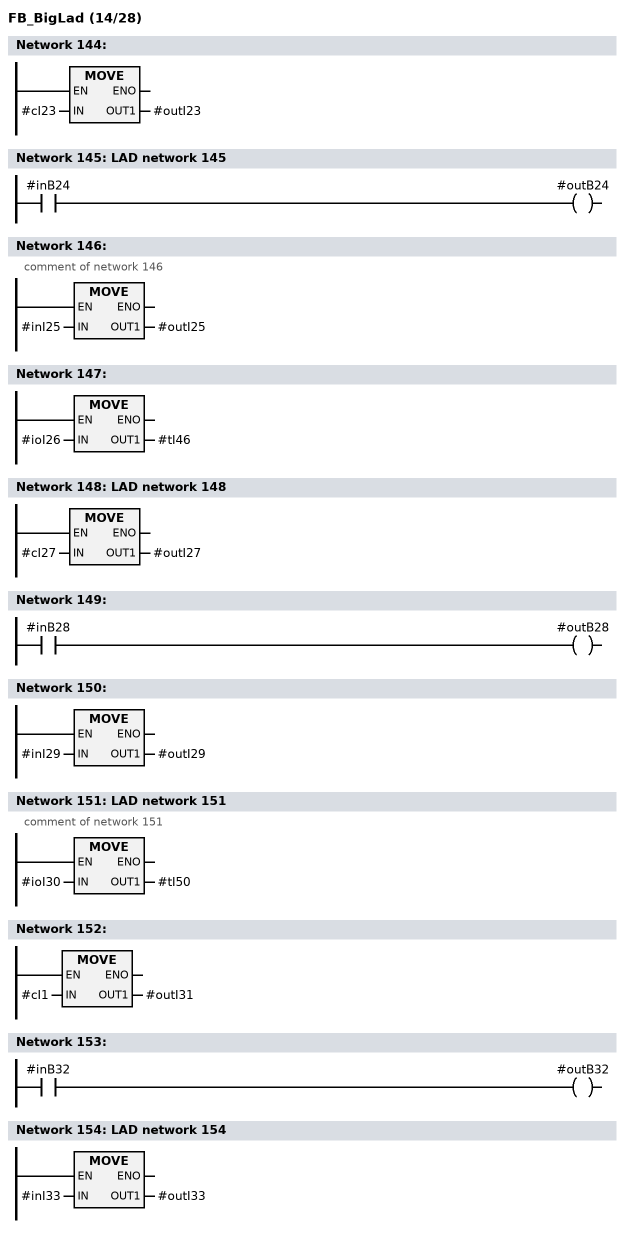
   RUNG wire#powerrail
      Move(in := #cI23, out1 => #outI23)
   END_RUNG
   // the same network as SCL:
   #outI23 := #cI23;
END_REGION

REGION Network 145: LAD network 145
   RUNG wire#powerrail
      Contact( #inB24 )
      Coil( #outB24 )
   END_RUNG
   // the same network as SCL:
   #outB24 := #inB24;
END_REGION

REGION Network 146
   // comment of network 146
   RUNG wire#powerrail
      Move(in := #inI25, out1 => #outI25)
   END_RUNG
   // the same network as SCL:
   #outI25 := #inI25;
END_REGION

REGION Network 147
   RUNG wire#powerrail
      Move(in := #ioI26, out1 => #tI46)
   END_RUNG
   // the same network as SCL:
   #tI46 := #ioI26;
END_REGION

REGION Network 148: LAD network 148
   RUNG wire#powerrail
      Move(in := #cI27, out1 => #outI27)
   END_RUNG
   // the same network as SCL:
   #outI27 := #cI27;
END_REGION

REGION Network 149
   RUNG wire#powerrail
      Contact( #inB28 )
      Coil( #outB28 )
   END_RUNG
   // the same network as SCL:
   #outB28 := #inB28;
END_REGION

REGION Network 150
   RUNG wire#powerrail
      Move(in := #inI29, out1 => #outI29)
   END_RUNG
   // the same network as SCL:
   #outI29 := #inI29;
END_REGION

REGION Network 151: LAD network 151
   // comment of network 151
   RUNG wire#powerrail
      Move(in := #ioI30, out1 => #tI50)
   END_RUNG
   // the same network as SCL:
   #tI50 := #ioI30;
END_REGION

REGION Network 152
   RUNG wire#powerrail
      Move(in := #cI1, out1 => #outI31)
   END_RUNG
   // the same network as SCL:
   #outI31 := #cI1;
END_REGION

REGION Network 153
   RUNG wire#powerrail
      Contact( #inB32 )
      Coil( #outB32 )
   END_RUNG
   // the same network as SCL:
   #outB32 := #inB32;
END_REGION

REGION Network 154: LAD network 154
   RUNG wire#powerrail
      Move(in := #inI33, out1 => #outI33)
   END_RUNG
   // the same network as SCL:
   #outI33 := #inI33;
END_REGION

REGION Network 155
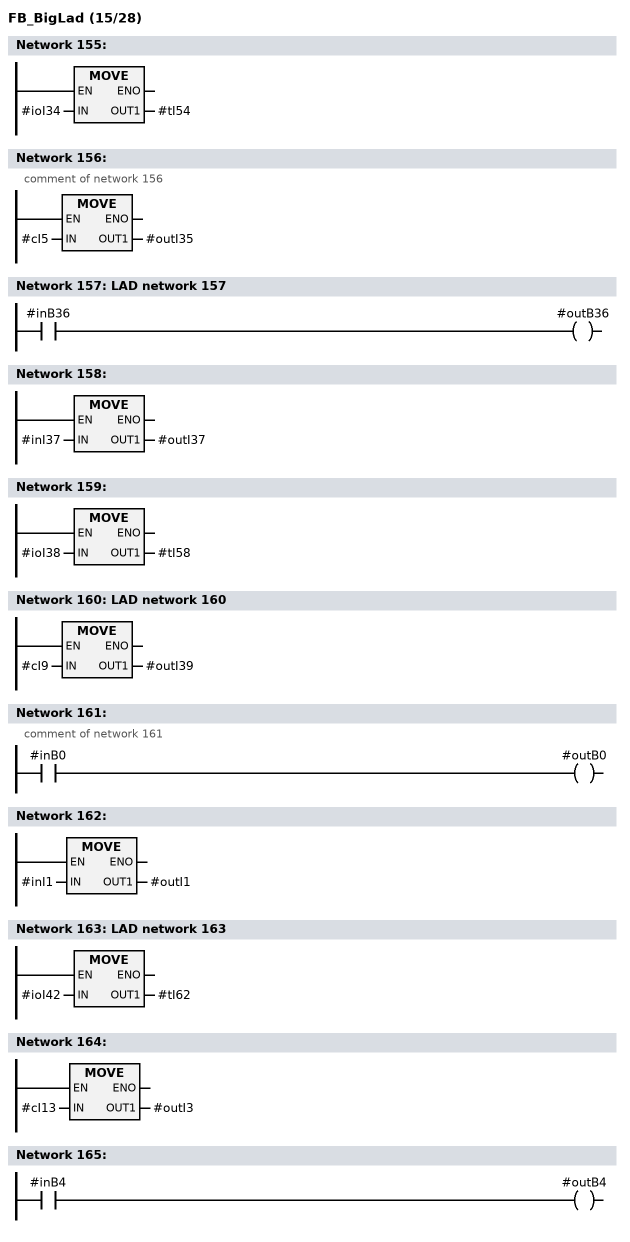
   RUNG wire#powerrail
      Move(in := #ioI34, out1 => #tI54)
   END_RUNG
   // the same network as SCL:
   #tI54 := #ioI34;
END_REGION

REGION Network 156
   // comment of network 156
   RUNG wire#powerrail
      Move(in := #cI5, out1 => #outI35)
   END_RUNG
   // the same network as SCL:
   #outI35 := #cI5;
END_REGION

REGION Network 157: LAD network 157
   RUNG wire#powerrail
      Contact( #inB36 )
      Coil( #outB36 )
   END_RUNG
   // the same network as SCL:
   #outB36 := #inB36;
END_REGION

REGION Network 158
   RUNG wire#powerrail
      Move(in := #inI37, out1 => #outI37)
   END_RUNG
   // the same network as SCL:
   #outI37 := #inI37;
END_REGION

REGION Network 159
   RUNG wire#powerrail
      Move(in := #ioI38, out1 => #tI58)
   END_RUNG
   // the same network as SCL:
   #tI58 := #ioI38;
END_REGION

REGION Network 160: LAD network 160
   RUNG wire#powerrail
      Move(in := #cI9, out1 => #outI39)
   END_RUNG
   // the same network as SCL:
   #outI39 := #cI9;
END_REGION

REGION Network 161
   // comment of network 161
   RUNG wire#powerrail
      Contact( #inB0 )
      Coil( #outB0 )
   END_RUNG
   // the same network as SCL:
   #outB0 := #inB0;
END_REGION

REGION Network 162
   RUNG wire#powerrail
      Move(in := #inI1, out1 => #outI1)
   END_RUNG
   // the same network as SCL:
   #outI1 := #inI1;
END_REGION

REGION Network 163: LAD network 163
   RUNG wire#powerrail
      Move(in := #ioI42, out1 => #tI62)
   END_RUNG
   // the same network as SCL:
   #tI62 := #ioI42;
END_REGION

REGION Network 164
   RUNG wire#powerrail
      Move(in := #cI13, out1 => #outI3)
   END_RUNG
   // the same network as SCL:
   #outI3 := #cI13;
END_REGION

REGION Network 165
   RUNG wire#powerrail
      Contact( #inB4 )
      Coil( #outB4 )
   END_RUNG
   // the same network as SCL:
   #outB4 := #inB4;
END_REGION

REGION Network 166: LAD network 166
   // comment of network 166
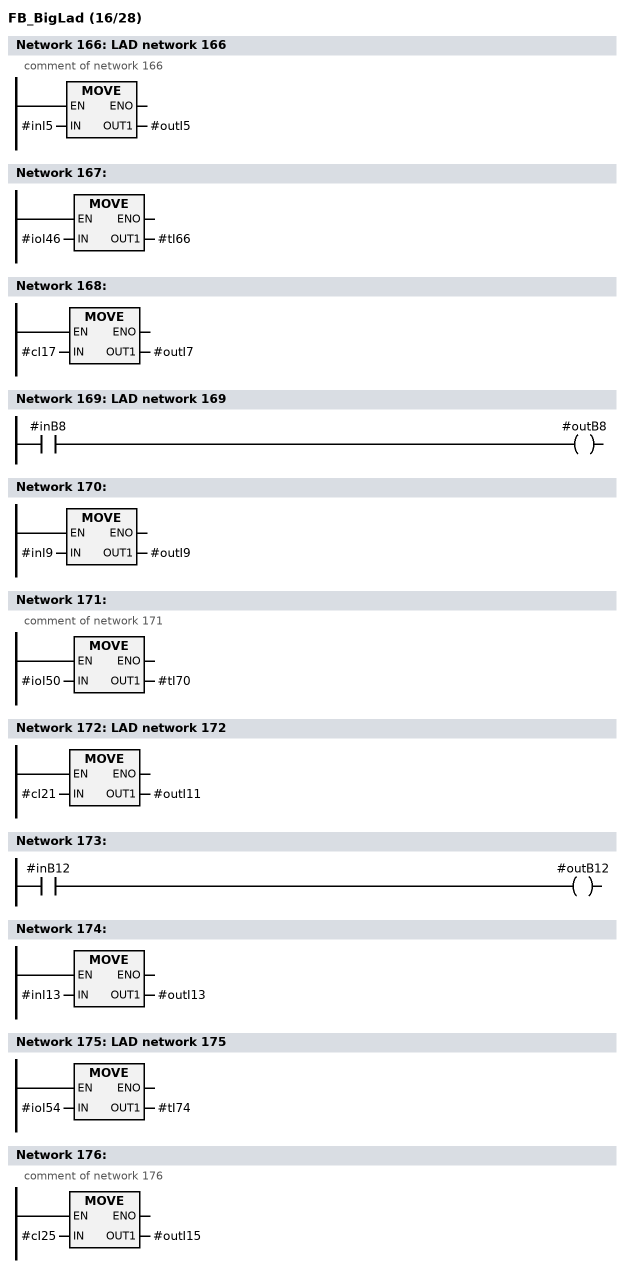
   RUNG wire#powerrail
      Move(in := #inI5, out1 => #outI5)
   END_RUNG
   // the same network as SCL:
   #outI5 := #inI5;
END_REGION

REGION Network 167
   RUNG wire#powerrail
      Move(in := #ioI46, out1 => #tI66)
   END_RUNG
   // the same network as SCL:
   #tI66 := #ioI46;
END_REGION

REGION Network 168
   RUNG wire#powerrail
      Move(in := #cI17, out1 => #outI7)
   END_RUNG
   // the same network as SCL:
   #outI7 := #cI17;
END_REGION

REGION Network 169: LAD network 169
   RUNG wire#powerrail
      Contact( #inB8 )
      Coil( #outB8 )
   END_RUNG
   // the same network as SCL:
   #outB8 := #inB8;
END_REGION

REGION Network 170
   RUNG wire#powerrail
      Move(in := #inI9, out1 => #outI9)
   END_RUNG
   // the same network as SCL:
   #outI9 := #inI9;
END_REGION

REGION Network 171
   // comment of network 171
   RUNG wire#powerrail
      Move(in := #ioI50, out1 => #tI70)
   END_RUNG
   // the same network as SCL:
   #tI70 := #ioI50;
END_REGION

REGION Network 172: LAD network 172
   RUNG wire#powerrail
      Move(in := #cI21, out1 => #outI11)
   END_RUNG
   // the same network as SCL:
   #outI11 := #cI21;
END_REGION

REGION Network 173
   RUNG wire#powerrail
      Contact( #inB12 )
      Coil( #outB12 )
   END_RUNG
   // the same network as SCL:
   #outB12 := #inB12;
END_REGION

REGION Network 174
   RUNG wire#powerrail
      Move(in := #inI13, out1 => #outI13)
   END_RUNG
   // the same network as SCL:
   #outI13 := #inI13;
END_REGION

REGION Network 175: LAD network 175
   RUNG wire#powerrail
      Move(in := #ioI54, out1 => #tI74)
   END_RUNG
   // the same network as SCL:
   #tI74 := #ioI54;
END_REGION

REGION Network 176
   // comment of network 176
   RUNG wire#powerrail
      Move(in := #cI25, out1 => #outI15)
   END_RUNG
   // the same network as SCL:
   #outI15 := #cI25;
END_REGION

REGION Network 177
